TYPE ST_PolarIIChamber_SelectThreeServiceStatus :
STRUCT
	Select1 : ST_ServiceStatus;
	Select2 : ST_ServiceStatus;
	Select3 : ST_ServiceStatus;
END_STRUCT
END_TYPE

(* stored: Version 1.1.0.1, ProductVersion 3.1.4026.18
   DUT ST_PolarIIChamber_SelectThreeServiceStatus: Id {14000000-0000-0000-0000-000000000042} *)
